Fanuc KAREL source: KO00141.KL

PROGRAM KO00141
%NOLOCKGROUP
VAR
  R: REAL
  CFG: CONFIG
  OUT: XYZWPR
  N: INTEGER
BEGIN
  N = 1
  R = 2.0
  CFG.CFG_FLIP = TRUE
  OUT = POS(R, R, R, N, R, R, CFG)
END KO00141
